Fanuc KAREL source: KO00102.KL

PROGRAM KO00102
%NOLOCKGROUP
VAR
  A: INTEGER
  B: ARRAY[2] OF BYTE
  OUT: REAL
BEGIN
  A = 1
  B[1] = 2
  OUT = ATAN2(A, B[1])
END KO00102
